(* IEC 61131-3 sources: openplc-editor-canopen/src/backend/shared/transpilers/st-transpiler/__tests__/fixtures/ld-relayout-corpus/ld-corpus-parallel-width/expected-st, 3 files *)

(* ---- _project.st ---- *)
CONFIGURATION Config0

  RESOURCE Res0 ON PLC
    TASK task0(INTERVAL := T#20ms,PRIORITY := 1);
    PROGRAM instance0 WITH task0 : main;
  END_RESOURCE
END_CONFIGURATION

(* ---- Blocks.st ---- *)
PROGRAM Blocks
  VAR
    TON0 : TON;
    w06_y : BOOL;
    w06_b : BOOL;
    w06_a : BOOL;
    w07_c : BOOL;
    CTU0 : CTU;
    w07_y : BOOL;
    w07_i : BOOL;
    w07_k : BOOL;
    w07_j : BOOL;
    w08_c : BOOL;
    CTUD0 : CTUD;
    w08_y : BOOL;
    w08_i : BOOL;
    w08_k : BOOL;
    w08_l : BOOL;
    w08_j : BOOL;
  END_VAR

  TON0(IN := w06_a, PT := T#1s);
  w06_y := TON0.Q OR w06_b;
  CTU0(CU := w07_c, R := w07_k OR w07_j AND w07_i);
  w07_y := CTU0.Q;
  CTUD0(CU := w08_c, LD := w08_k OR w08_l OR w08_j AND w08_i);
  w08_y := CTUD0.QU;
END_PROGRAM

(* ---- Branches.st ---- *)
PROGRAM Branches
  VAR
    w01_a : BOOL;
    w01_y : BOOL;
    w01_b : BOOL;
    w01_e : BOOL;
    w01_c : BOOL;
    w01_d : BOOL;
    w02_f : BOOL;
    w02_y : BOOL;
    w02_g : BOOL;
    w02_j : BOOL;
    w02_h : BOOL;
    w02_i : BOOL;
    w02_k : BOOL;
    w03_e : BOOL;
    w03_y : BOOL;
    w03_a : BOOL;
    w03_b : BOOL;
    w03_d : BOOL;
    w03_c : BOOL;
    w04_a : BOOL;
    w04_y : BOOL;
    w04_conveyor_infeed_photoeye_blocked_longer_than_limit : BOOL;
    w04_b : BOOL;
    w05_a : BOOL;
    w05_k : BOOL;
    w05_conveyor_reject_gate_solenoid_output_main : BOOL;
  END_VAR

  w01_y := (w01_e OR w01_d AND w01_c AND w01_b) AND w01_a;
  w02_y := w02_f OR w02_i AND w02_h AND w02_g OR w02_k AND w02_j;
  w03_y := w03_e OR (w03_d OR w03_c AND w03_b) AND w03_a;
  w04_y := w04_conveyor_infeed_photoeye_blocked_longer_than_limit OR w04_b AND w04_a;
  w05_k := w05_a;
  w05_conveyor_reject_gate_solenoid_output_main := w05_a;
END_PROGRAM
